(* IEC 61131-3 sources: TetherPLC/tests/ld, 5 files *)

(* ---- 01_start_hold_stop.st ---- *)
PROGRAM LD01_START_HOLD_STOP
VAR
    start_in AT %IX0.0 : BOOL;
    hold_in  AT %IX0.1 : BOOL;
    stop_in  AT %IX0.2 : BOOL;
    run_out  AT %QX0.0 : BOOL;
    lamp_out AT %QX0.1 : BOOL;
END_VAR
run_out := start_in AND hold_in AND NOT stop_in;
lamp_out := run_out;
END_PROGRAM

(* ---- 02_multi_coil.st ---- *)
PROGRAM LD02_MULTI_COIL
VAR
    a_in  AT %IX0.0 : BOOL;
    b_in  AT %IX0.1 : BOOL;
    c_out AT %QX0.0 : BOOL;
    d_out AT %QX0.1 : BOOL;
    e_out AT %QX0.2 : BOOL;
END_VAR
c_out := a_in AND b_in;
d_out := a_in AND b_in;
e_out := NOT a_in;
END_PROGRAM

(* ---- 03_parallel.st ---- *)
PROGRAM LD03_PARALLEL
VAR
    start_in AT %IX0.0 : BOOL;
    hold_in  AT %IX0.1 : BOOL;
    stop_in  AT %IX0.2 : BOOL;
    run_out  AT %QX0.0 : BOOL;
END_VAR
run_out := (start_in OR hold_in) AND NOT stop_in;
END_PROGRAM

(* ---- 04_fb_op.st ---- *)
PROGRAM P04_LD_FB_OP
VAR
    start_in AT %IX0.0 : BOOL;
    stop_in AT %IX0.1 : BOOL;
    run AT %QX0.0 : BOOL;
    ton1 : TON;
END_VAR
ton1(IN := start_in, PT := T#200ms);
run := ton1.Q AND NOT stop_in;
END_PROGRAM

(* ---- 05_data.st ---- *)
PROGRAM P05_LD_DATA
VAR
    a AT %IX0.0 : BOOL;
    b AT %IX0.1 : BOOL;
    c AT %IX0.2 : BOOL;
    t AT %MX0.0 : BOOL;
    y AT %QX0.0 : BOOL;
END_VAR
t := a AND b;
y := t OR c;
END_PROGRAM
